// TwinCAT 3 PLC project Untitled1
// ProgramVersion: 3.1.4026.26
// libraries:
//   Tc2_Standard, * (Beckhoff Automation GmbH)
//   Tc2_System, * (Beckhoff Automation GmbH)
// project tree:
//   DUTs/ coffee.TcDUT, tea.TcDUT
//   GVLs/ gvl.TcGVL
//   / PlcTask.TcTTO
//   POUs/ MAIN.TcPOU
// real-time tasks:
//   TASK PlcTask: cycle T#10ms, priority 20, ADS port 350

CONFIGURATION Untitled1
    RESOURCE PLC ON TwinCAT3
        TASK PlcTask(INTERVAL := T#10ms, PRIORITY := 20);
        PROGRAM MAIN WITH PlcTask : MAIN;
    END_RESOURCE
END_CONFIGURATION

// ---- DUTs/coffee.TcDUT
TYPE coffee :
STRUCT
	
price			: REAL;
name			: STRING;
ingredients		: STRING;


END_STRUCT
END_TYPE

// ---- DUTs/tea.TcDUT
TYPE tea :
STRUCT

price			: REAL;
name			: STRING;
ingredients		: STRING;	


END_STRUCT
END_TYPE

// ---- GVLs/gvl.TcGVL
{attribute 'qualified_only'}
VAR_GLOBAL
	
coffees			: coffee;
teas			: tea;

END_VAR

// ---- POUs/MAIN.TcPOU
PROGRAM MAIN
VAR
	
tempVar			: BOOL;

END_VAR

END_PROGRAM
